Yaskawa INFORM job: UTEST10.JBI

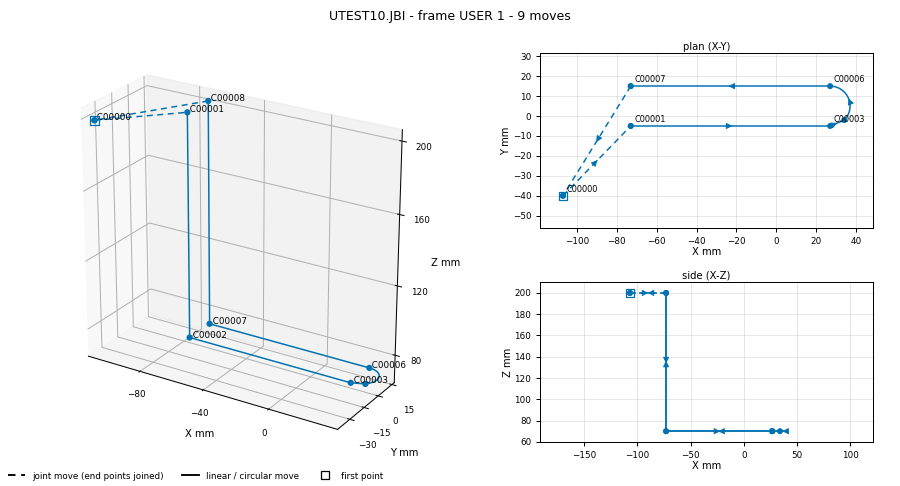
[picture p0: tool path of UTEST10.JBI in frame USER 1, 9 of 10 moves have a stored position in this frame; points joined in program order, loops and branches not executed]
/JOB
//NAME UTEST10
//POS
///NPOS 10,0,0,0,0,0
///USER 1
///TOOL 1
///POSTYPE USER
///RECTAN
///RCONF 1,0,0,0,0,0,0,0,0,0,0,0,0,0,0,0,0,0,0,0,0,0,0,0
C00000=-107.000,-40.000,200.000,0.0000,0.0000,-150.0000
C00001=-73.000,-5.000,200.000,0.0000,0.0000,-150.0000
C00002=-73.000,-5.000,70.000,0.0000,0.0000,-150.0000
C00003=27.000,-5.000,70.000,0.0000,0.0000,-150.0000
C00004=34.070,-2.070,70.000,0.0000,0.0000,-150.0000
C00005=34.070,12.070,70.000,0.0000,0.0000,-150.0000
C00006=27.000,15.000,70.000,0.0000,0.0000,-150.0000
C00007=-73.000,15.000,70.000,0.0000,0.0000,-150.0000
C00008=-73.000,15.000,200.000,0.0000,0.0000,-150.0000
C00009=-107.000,-40.000,200.000,0.0000,0.0000,-150.0000
//INST
///DATE 2026/11/25 16:27
///ATTR SC,RW,RJ
////FRAME USER 1
///GROUP1 RB1
NOP
MOVJ C00000 VJ=0.78
MOVJ C00001 VJ=0.78
MOVL C00002 V=11.0
MOVL C00003 V=10.0 ACC=20 DEC=20
MOVC C00004 V=12.0 ACC=20 DEC=20
MOVC C00005 V=12.0 ACC=20 DEC=20
MOVC C00006 V=12.0 ACC=20 DEC=20
MOVL C00007 V=10.0 ACC=20 DEC=20
MOVL C00008 V=11.0
MOVJ C00009 VJ=0.78
END
